(* PLC project constructs-0201-app.project, CODESYS CODESYS V3.5 SP17 Patch 3 *)
(* stored: creationDateTime 2026-10-19T09:47:53.8582923, modificationDateTime 1601-01-01T03:00:00 *)

// Перечисление без значений и без базового типа
TYPE E_Color :
(
    Red,
    Green,
    Blue
);
END_TYPE

// Режим устройства: перечисление с явными значениями и базовым типом
{attribute 'qualified_only'}
{attribute 'strict'}
TYPE E_Mode :
(
    OutOfService := 0,  // выведено из работы
    Auto := 1,          // автоматический
    Manual := 2,        // ручной
    Local := 3          // местный
) INT;
END_TYPE

// Базовая структура: начальные значения, массив, строка, комментарии
TYPE ST_Base :
STRUCT
    xEnable : BOOL := TRUE;               // разрешение
    iCount : INT;                         (* счётчик *)
    rValue_bar : REAL := 1.5;
    sName : STRING(32) := 'base';
    wsLabel : WSTRING(16) := "Насос";
    aiData : ARRAY[0..3] OF INT := [1, 2, 3, 4];
    eMode : E_Mode := E_Mode.Auto;
END_STRUCT
END_TYPE

// Структура-наследник базовой
TYPE ST_Derived EXTENDS ST_Base :
STRUCT
    tDelay : TIME := T#5S;
    ltStamp : LTIME;
    pData : POINTER TO INT;
END_STRUCT
END_TYPE

// Псевдоним строкового типа
TYPE T_Name : STRING(20);
END_TYPE

// Псевдоним с поддиапазоном
TYPE T_Percent : INT(0..100);
END_TYPE

// Команды двигателя от HMI (DUT в папке проекта)
TYPE ST_MotorCmd :
STRUCT
    xStart : BOOL;
    xStop : BOOL;
    eMode : E_Mode := E_Mode.OutOfService;
END_STRUCT
END_TYPE

// Состояние двигателя для HMI (DUT во вложенной папке Motor/Status)
TYPE ST_MotorSts :
STRUCT
    xRun : BOOL;
    uiStarts : UINT;
    eMode : E_Mode := E_Mode.OutOfService;
END_STRUCT
END_TYPE

// Устройство: режим, отказ, пуск
INTERFACE I_Device EXTENDS I_Resettable
METHOD Start : BOOL
END_METHOD
PROPERTY Fault : BOOL
END_PROPERTY
PROPERTY Mode : E_Mode
END_PROPERTY
END_INTERFACE

// Блокировка по месту
INTERFACE I_Lockable
METHOD Lock
VAR_INPUT
    xLock : BOOL;
END_VAR
END_METHOD
END_INTERFACE

// Позиционер: уставка (только запись) и перемещение
INTERFACE I_Positioner
// Переместить в позицию, %
METHOD MoveTo : BOOL
VAR_INPUT
    rPos_pct : REAL;
END_VAR
VAR_OUTPUT
    xDone : BOOL;
END_VAR
END_METHOD
PROPERTY Setpoint : REAL
END_PROPERTY
END_INTERFACE

// Сброс состояния
INTERFACE I_Resettable
// Сбросить; TRUE — сброс выполнен
METHOD Reset : BOOL
VAR_INPUT
    xForce : BOOL;
END_VAR
END_METHOD
END_INTERFACE

TYPE U_Raw : UNION
  wWord : WORD;
  aBytes : ARRAY[0..1] OF BYTE;
END_UNION;
END_TYPE

// Назначение: ограничение значения диапазоном [rMin, rMax]; при rMin > rMax границы меняются местами
// Автор:      <ИМЯ ФАМИЛИЯ>
// Версия:     0.1.0
// Документ:   docs/plcopen.md
FUNCTION F_Clamp : REAL
VAR_INPUT
    rValue : REAL;      // значение
    rMin : REAL;        // нижняя граница
    rMax : REAL;        // верхняя граница
END_VAR
VAR
    rLow : REAL;
    rHigh : REAL;
END_VAR

                  // границы в правильном порядке
IF rMin <= rMax THEN
    rLow := rMin;
    rHigh := rMax;
ELSE
    rLow := rMax;
    rHigh := rMin;
END_IF
F_Clamp := LIMIT(rLow, rValue, rHigh);

                
END_FUNCTION

// Назначение: функция без типа результата
// Автор:      <ИМЯ ФАМИЛИЯ>
// Версия:     0.1.0
// Документ:   docs/plcopen.md
FUNCTION F_Noop
VAR_INPUT
    xIn : BOOL;
END_VAR

                  // тела нет
;

                
END_FUNCTION

// Назначение: сумма элементов массива любой длины (VAR_IN_OUT CONSTANT, ARRAY[*])
// Автор:      <ИМЯ ФАМИЛИЯ>
// Версия:     0.1.0
// Документ:   docs/plcopen.md
FUNCTION F_Sum : LREAL
VAR_IN_OUT CONSTANT
    arValues : ARRAY[*] OF REAL;
END_VAR
VAR
    diIdx : DINT;
END_VAR

                  F_Sum := 0;
FOR diIdx := LOWER_BOUND(arValues, 1) TO UPPER_BOUND(arValues, 1) DO
    F_Sum := F_Sum + arValues[diIdx];
END_FOR

                
END_FUNCTION

// Назначение: счётчик фронтов с задержкой подтверждения (без ООП, Standard: R_TRIG, TON)
// Автор:      <ИМЯ ФАМИЛИЯ>
// Версия:     0.1.0
// Документ:   docs/plcopen.md
FUNCTION_BLOCK FB_Counter
VAR_INPUT
    xIn : BOOL;                 // вход
    tConfirm : TIME := T#100MS; // задержка подтверждения
END_VAR
VAR_OUTPUT
    udiCount : UDINT;           // число фронтов
    xConfirmed : BOOL;
END_VAR
VAR_IN_OUT
    stCmd : ST_MotorCmd;
END_VAR
VAR
    fbEdge : R_TRIG;
    fbDelay : TON;
END_VAR
VAR RETAIN
    udiTotal : UDINT;
END_VAR
VAR_TEMP
    xEdge : BOOL;
END_VAR

                  fbEdge(CLK := xIn);
xEdge := fbEdge.Q;
IF xEdge THEN
    udiCount := udiCount + 1;
    udiTotal := udiTotal + 1;
END_IF
fbDelay(IN := xIn, PT := tConfirm, Q => xConfirmed);
stCmd.xStart S= xConfirmed;
stCmd.xStop R= xConfirmed;

                
END_FUNCTION_BLOCK

// Назначение: программа с методом; комментарии всех видов
// Автор:      <ИМЯ ФАМИЛИЯ>
// Версия:     0.1.0
// Документ:   docs/plcopen.md
PROGRAM PRG_Aux
VAR
    fbValve : FB_Valve;
    itfPos : I_Positioner;
    itfLock : I_Lockable;
    iCalls : INT;
    wsMsg : WSTRING(32) := "Задвижка <закрыта> & 'ok'";
    sMsg : STRING(32) := 'a$'b"c <&>';
END_VAR
VAR_EXTERNAL
    xDoRun : BOOL;              // выход из GVL_Io (необязательное объявление CODESYS)
END_VAR

                  (* внешний (* вложенный *) комментарий *)
itfPos := fbValve;
itfLock := fbValve;
itfPos.Setpoint := 50.0;
itfPos.MoveTo(rPos_pct := 40.0);
itfLock.Lock(xLock := NOT xDoRun);
fbValve();
Step(iInc := 1);
F_Noop(xIn := TRUE);
IF iCalls > 5 AND_THEN fbValve.rPos_pct < 1.0E3 THEN
    iCalls := 0;
END_IF

                

// Шаг программы
METHOD Step : INT
VAR_INPUT
    iInc : INT := 1;
END_VAR
                        iCalls := iCalls + iInc;
Step := iCalls;

                      
END_METHOD
END_PROGRAM

// Назначение: точка входа — вызывает все объекты примера
// Автор:      <ИМЯ ФАМИЛИЯ>
// Версия:     0.1.0
// Документ:   docs/plcopen.md
PROGRAM PRG_Main
VAR
    fbMotor : FB_Motor;
    itfDevice : I_Device;
    itfReset : I_Resettable;
    fbCounter : FB_Counter;
    stCmd : ST_MotorCmd;
    stSts : ST_MotorSts;
    stDerived : ST_Derived;
    uRaw : U_Raw;
    ePercent : T_Percent := 50;
    sName : T_Name := 'pump';
    eColor : E_Color := E_Color.Green;
    arBuf : ARRAY[0..2] OF REAL := [3(1.0)];
    rOut : REAL;
    lrSum : LREAL;
    pValue : POINTER TO REAL;
    refValue : REFERENCE TO REAL;
    iStep : INT;
    xOk : BOOL;
END_VAR

                  (* вызовы всех объектов примера *)
itfDevice := fbMotor;
itfReset := fbMotor;
fbMotor(stCmd := stCmd);
IF itfDevice <> 0 THEN
    itfDevice.Mode := E_Mode.Auto;
    xOk := itfDevice.Fault;
END_IF
itfReset.Reset(xForce := TRUE);
fbCounter(xIn := GVL_Io.xDiStart, stCmd := GVL_Io.astCmd[GVL_Io.IO_CHANNELS - 1]);
GVL_Io.xDoRun := fbMotor.xRun;
stSts.xRun := fbMotor.xRun;
stSts.uiStarts := fbMotor.Starts;
rOut := F_Clamp(rValue := INT_TO_REAL(GVL_Io.iAiLevel), rMin := 0.0, rMax := 100.0);
lrSum := F_Sum(arValues := arBuf);
pValue := ADR(rOut);
refValue REF= rOut;
IF __ISVALIDREF(refValue) THEN
    refValue := refValue + GVL_Const.RATE_LIMIT;
END_IF
uRaw.wWord := 16#1234;
stDerived.tDelay := T#1S;
CASE iStep OF
    0:
        iStep := 1;
    1, 2:
        iStep := iStep + 1;
ELSE
    iStep := 0;
END_CASE
WHILE iStep > 10 DO
    iStep := iStep - 1;
END_WHILE
REPEAT
    iStep := iStep + 0;
UNTIL TRUE
END_REPEAT
GVL_Io.udiRunHours := GVL_Io.udiRunHours + fbCounter.udiCount;
PersistentVars.udiStartsTotal := PersistentVars.udiStartsTotal + fbMotor.Starts;
sName := GVL_Const.TEXT_OK;
eColor := E_Color.Blue;
ePercent := 75;
PRG_Aux();

                
END_PROGRAM

// Назначение: абстрактная база устройств — режим, отказ, квитирование
// Автор:      <ИМЯ ФАМИЛИЯ>
// Версия:     0.1.0
// Документ:   docs/plcopen.md
{attribute 'reflection'}
FUNCTION_BLOCK ABSTRACT FB_DeviceBase IMPLEMENTS I_Device
VAR_INPUT
    xReset : BOOL;
END_VAR
VAR_OUTPUT
    xFault : BOOL;
END_VAR
VAR
    eModeInt : E_Mode := E_Mode.OutOfService;
    {attribute 'hide'}
    xFaultInt : BOOL;
END_VAR
VAR_STAT
    uiInstances : UINT;
END_VAR

                  // общая логика базы: сброс по входу
IF xReset THEN
    Reset(xForce := FALSE);
END_IF
xFault := xFaultInt;

                

// Сброс отказа
METHOD PUBLIC Reset : BOOL
VAR_INPUT
    xForce : BOOL;
END_VAR
                        xFaultInt := FALSE;
Reset := TRUE;

                      
END_METHOD

// Установить отказ (только для наследников)
METHOD PROTECTED SetFault
VAR_INPUT
    xValue : BOOL;
END_VAR
                        xFaultInt := xValue;

                      
END_METHOD

// Пуск — реализует наследник
METHOD PUBLIC ABSTRACT Start : BOOL
                        
                      
END_METHOD

PROPERTY PUBLIC Fault : BOOL
GET
VAR
END_VAR
                          Fault := xFaultInt;

                        
END_GET
END_PROPERTY

// Текущий режим
PROPERTY PUBLIC Mode : E_Mode
GET
VAR
END_VAR
                          Mode := eModeInt;

                        
END_GET
SET
VAR
END_VAR
                          eModeInt := Mode;

                        
END_SET
END_PROPERTY
END_FUNCTION_BLOCK

// Назначение: двигатель — наследник базы: пуск, сброс через SUPER^, счёт пусков
// Автор:      <ИМЯ ФАМИЛИЯ>
// Версия:     0.1.0
// Документ:   docs/plcopen.md
FUNCTION_BLOCK FB_Motor EXTENDS FB_DeviceBase
VAR_INPUT
    stCmd : ST_MotorCmd;
END_VAR
VAR_OUTPUT
    xRun : BOOL;
END_VAR
VAR
    uiStarts : UINT;
    fbCounter : FB_Counter;
END_VAR

                  SUPER^();
IF stCmd.xStart AND NOT xFault THEN
    Start();
ELSIF stCmd.xStop THEN
    xRun := FALSE;
END_IF

                

// Описание для журнала
METHOD PRIVATE FINAL Describe : WSTRING(40)
VAR
    wsText : WSTRING(40) := "Двигатель";
END_VAR
                        Describe := wsText;

                      
END_METHOD

// Инициализация экземпляра
METHOD FB_init : BOOL
VAR_INPUT
    bInitRetains : BOOL;    // TRUE — инициализировать RETAIN
    bInCopyCode : BOOL;     // TRUE — экземпляр копируется при онлайн-изменении
END_VAR
                        uiStarts := 0;

                      
END_METHOD

METHOD PUBLIC Reset : BOOL
VAR_INPUT
    xForce : BOOL;
END_VAR
                        Reset := SUPER^.Reset(xForce := xForce);
xRun := FALSE;

                      
END_METHOD

METHOD PUBLIC Start : BOOL
VAR_INST
    uiCalls : UINT;     // число вызовов метода (сохраняется между вызовами)
END_VAR
                        uiCalls := uiCalls + 1;
IF THIS^.Mode = E_Mode.Auto OR Mode = E_Mode.Manual THEN
    xRun := TRUE;
    uiStarts := uiStarts + 1;
END_IF
Start := xRun;

                      
END_METHOD

// Число пусков
PROPERTY PUBLIC Starts : UINT
GET
VAR
    uiCopy : UINT;
END_VAR
                          uiCopy := uiStarts;
Starts := uiCopy;

                        
END_GET
SET
VAR
END_VAR
                          uiStarts := Starts;

                        
END_SET
END_PROPERTY
END_FUNCTION_BLOCK

// Назначение: задвижка — FINAL-наследник базы с двумя интерфейсами
// Автор:      <ИМЯ ФАМИЛИЯ>
// Версия:     0.1.0
// Документ:   docs/plcopen.md
FUNCTION_BLOCK FINAL FB_Valve EXTENDS FB_DeviceBase IMPLEMENTS I_Positioner, I_Lockable
VAR_OUTPUT
    rPos_pct : REAL;
    xLocked : BOOL;
END_VAR
VAR
    rSetpoint_pct : REAL;
END_VAR
VAR CONSTANT
    POS_MAX : REAL := 100.0;
END_VAR

                  SUPER^();
IF NOT xLocked THEN
    rPos_pct := F_Clamp(rValue := rSetpoint_pct, rMin := 0.0, rMax := POS_MAX);
END_IF

                

METHOD PUBLIC Lock
VAR_INPUT
    xLock : BOOL;
END_VAR
                        xLocked := xLock;

                      
END_METHOD

METHOD PUBLIC MoveTo : BOOL
VAR_INPUT
    rPos_pct : REAL;
END_VAR
VAR_OUTPUT
    xDone : BOOL;
END_VAR
                        rSetpoint_pct := rPos_pct;
xDone := THIS^.rPos_pct = rPos_pct;
MoveTo := NOT xLocked;

                      
END_METHOD

METHOD PUBLIC Start : BOOL
                        Start := NOT xLocked;

                      
END_METHOD

// Внутренний метод библиотеки
METHOD INTERNAL Trace : ST_MotorCmd
VAR_IN_OUT
    stLast : ST_MotorCmd;
END_VAR
                        Trace := stLast;

                      
END_METHOD

PROPERTY PUBLIC Setpoint : REAL
SET
VAR
END_VAR
                          rSetpoint_pct := Setpoint;

                        
END_SET
END_PROPERTY
END_FUNCTION_BLOCK

CONFIGURATION Application
  RESOURCE Application ON PLC
(* global variable list GVL_Const *)
// Константы
{attribute 'qualified_only'}
VAR_GLOBAL CONSTANT
    MAX_ITEMS : INT := 4;           // число элементов
    RATE_LIMIT : REAL := 0.25;
    TEXT_OK : STRING := 'OK';
END_VAR
(* global variable list GVL_Io *)
// Входы-выходы и сохраняемые значения
VAR_GLOBAL
    xDiStart AT %IX0.0 : BOOL;      // кнопка «Пуск»
    xDoRun AT %QX0.0 : BOOL;
    iAiLevel AT %IW2 : INT;
    astCmd : ARRAY[1..GVL_Const.MAX_ITEMS] OF ST_MotorCmd;
END_VAR
VAR_GLOBAL RETAIN
    udiRunHours : UDINT;
END_VAR
VAR_GLOBAL CONSTANT
    IO_CHANNELS : INT := 2;         // число каналов (константа в одном списке с переменными)
END_VAR
(* global variable list PersistentVars *)
// Сохраняемые переменные (объект Persistent Variables)
VAR_GLOBAL PERSISTENT RETAIN
    udiStartsTotal : UDINT;     // пуски за весь срок службы
    rRunHours_h : REAL;
END_VAR
  END_RESOURCE
END_CONFIGURATION
